Fanuc KAREL source: kb00150.compact.KL

PROGRAM KB00150
%STACKSIZE=65535
%PRIORITY=65535
%NOLOCKGROUP
VAR
P1 : STRING[80]
P2 : STRING[80]
P3 : STRING[80]
P4 : STRING[80]
P5 : INTEGER
BEGIN
P1='A'
P2='A'
P3='A'
P4='A'
P5=1
RMCN_ALERT(P1,P2,P3,P4,P5)
END KB00150
